// SIMATIC S7-200 project (STEP 7-Micro/WIN), CPU 224 CN REL 02.01

SYMBOL_TABLE ????1
boton_sb1        I1.2
boton_sb2        I1.3
selector         I1.5
parada           I1.4
act1             Q0.0
act2             Q0.1
END_SYMBOL_TABLE

ORGANIZATION_BLOCK ???:OB1
TITLE=????
BEGIN
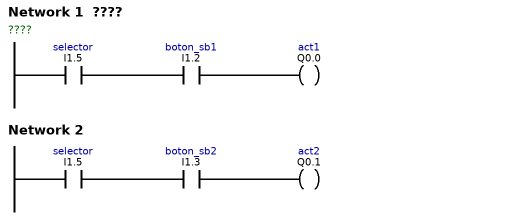
Network 1 // ????
// ????
LD     selector:I1.5
A      boton_sb1:I1.2
=      act1:Q0.0
Network 2
LD     selector:I1.5
A      boton_sb2:I1.3
=      act2:Q0.1
END_ORGANIZATION_BLOCK
